(* Logix 5000 project; controller TFF vendor 1 type 14 code 107 rev 34.11; software revision 34.03; part 13 of 36 *)
(* tags used below, declared in another part *)
   AlarmAnalog : AlarmAnalog[50];   // Analog Alarm Array
   AlarmControl : AlarmControl;   // Alarm Control
   AlarmDeviation : AlarmDeviation[20];   // Control Loop Deviation Alarm Array
   AnalogPoint : AnalogInput[50];   // Analog Input Array
   CCPSystem : CCPSystem;   // CCP System Data
   ChartMark : ChartMark;   // Chart Mark
   Concentration : Concentration;
   ControlLoop : ControlLoop[20];   // Control Loop Array
   CriteriaFlag : CriteriaFlag;   // Criteria Flag used in CCP Recipe
   DCS : DCS;
   DerivedData : DerivedData;   // Derived data (user input and calculated values)
   Diafiltration : Diafiltration;
   DigitalPoint : DigitalPoint[150];   // Digital Point Array
   Drive : Drive[11];   // Drives Array
   FlowPath : FlowPath[64];   // Flow Path Array
   FlowPathControl : FlowPathControl;   // Flow Path Control
   FQ_Conc : ALIAS FOR Totalizer[0];   // Concentration Totalizer
   FQ_Diaf : ALIAS FOR Totalizer[1];   // DiafiltrationTotalizer
   LogVal : LoggedValue;   // Setpoints to be logged
   Membrane_Data : Membrane_Data;   // Membrane Data
   MiscBOOL : BOOL[64];   // Misc BOOL Values
   MiscDINT : DINT[32];   // Misc DINT Values
   MiscREAL : REAL[50];   // Misc Real Values
   Mixer : Mixer;   // Mixer config. structure
   Operation : Operation[6,251];   // Operation Table
   PCV001_Control : PCV_Control;   // PCV001 Control UDT
   PCV101_Control : PCV_Control;   // PCV101 Control UDT
   Phase : Phases[6];   // Phase Control Array
   Phase0 : ALIAS FOR Phase[0];   // Phase 0
   Phase1 : ALIAS FOR Phase[1];   // Phase 1
   Phase2 : ALIAS FOR Phase[2];   // Phase 2
   Phase3 : ALIAS FOR Phase[3];   // Phase 3
   Phase4 : ALIAS FOR Phase[4];   // Phase 4
   Phase5 : ALIAS FOR Phase[5];   // Phase 5
   PhaseTotalizer : PhaseTotalizer[18];   // Phase Totalizers Array
   Prompt : Prompt[7];   // Prompt Array
   Prompt0 : ALIAS FOR Prompt[0];   // Phase 0 Prompt
   Prompt1 : ALIAS FOR Prompt[1];   // Phase 1 Prompt
   Prompt2 : ALIAS FOR Prompt[2];   // Phase 2 Prompt
   Prompt3 : ALIAS FOR Prompt[3];   // Phase 3 Prompt
   Prompt4 : ALIAS FOR Prompt[4];   // Phase 4 Prompt
   Prompt5 : ALIAS FOR Prompt[5];   // Phase 5 Prompt
   PromptTimer : FBD_TIMER;   // Prompt Timer
   SRL001 : ALIAS FOR DigitalPoint[15];   // Tank Skid Remote / Standalone
   SysControl : SysControl;   // General system status and command
   Tank : TankManagement;   // Tank Management
   ThisSystem : SystemType;
   Timers : Timers[22];   // Timer Array
   Totalizer : Totalizers[20];   // Totalizers Array
   UserAlarm : UserAlarm;   // User Alarm (used in CCP Recipe)
   UserTotalizerManagement : UserTotalizerManagement;   // User Totalizer management
   Valve : Valve[100];   // Valve Array
   Y500A : ALIAS FOR DigitalOutput[11];   // Unlock Clamshell
   Y500B : ALIAS FOR DigitalOutput[12];   // Lock Clamshell
   Y501A : ALIAS FOR DigitalOutput[10];   // Unlock Door
   Y501B : ALIAS FOR DigitalOutput[9];   // Lock Door
   Y502A : ALIAS FOR DigitalOutput[13];   // Unlock Clamshell in Door
   Y502B : ALIAS FOR DigitalOutput[14];   // Lock Clamshell in Door
   Y503A : ALIAS FOR DigitalOutput[15];   // Connect Clamshell
   Y503B : ALIAS FOR DigitalOutput[16];   // Disconnect Clamshell

PROGRAM CCPSystem   (* main routine MainRoutine, fault routine FaultRoutine *)
VAR
   ActionCode : DINT := 1700011;   // Action Code
   ActionFlag : BOOL;   // Action Flag
   ActionProperty : DINT := 11;   // Action Property
   ActionStructure : DINT := 17;   // Action Data Structure
   ActionTag : DINT;   // Action Tag
   ActionValue : REAL := 1.0;   // Action Value
   AutoRunTimer : TIMER := (PRE := 5000);   // Auto Run Timer
   Boolean : DINT;   // Boolean Operator
        .1   // AND
        .0   // OR
   Branch : BOOL;   // Conditional Branch Flag
   BranchStep : DINT;   // Branch Step Number
   BufferStep : DINT := 60;   // Buffer Step
   Clear : BOOL;   // Clear Operation Table Flag
   Code : DINT := 3100002;   // Global Code
   CompleteTimer : TIMER := (PRE := 10000);   // Operation Complete Timer
   Criteria1BoolValue : BOOL;   // Criteria 1 Discrete Value
   Criteria1Code : DINT := 1100602;   // Criteria 1 Code
   Criteria1Met : BOOL := 1;   // Criteria 1 Met
   Criteria1Operator : DINT := 1;   // Criteria 1 Operator
        .0   // >=
        .1   // <=
        .2   // =
   Criteria1Property : DINT := 2;   // Criteria 1 Property
   Criteria1RealValue : REAL := 2.0;   // Criteria 1 Real Value
   Criteria1Structure : DINT := 11;   // Criteria 1 Data Structure
   Criteria1Tag : DINT := 6;   // Criteria 1 Tag
   Criteria1Type : BOOL;   // Criteria 1 Type 0=Real, 1=Boolean
   Criteria1Value : REAL := 2.0;   // Criteria 1 Value
   Criteria2BoolValue : BOOL := 1;   // Criteria 2 Discrete Value
   Criteria2Code : DINT;   // Criteria 2 Code
   Criteria2Met : BOOL := 1;   // Criteria 2 Met
   Criteria2Operator : DINT;   // Criteria 2 Operator
        .0   // >=
        .1   // <=
        .2   // =
   Criteria2Property : DINT := 3;   // Criteria 2 Property
   Criteria2RealValue : REAL := 6.0;   // Criteria 2 Real Value
   Criteria2Structure : DINT;   // Criteria 2 Data Structure
   Criteria2Tag : DINT;   // Criteria 2 Tag
   Criteria2Type : BOOL;   // Criteria 2 Type 0=Real, 1=Boolean
   Criteria2Value : REAL;   // Criteria 2 Value
   CriteriaMet : BOOL := 1;   // Criteria Met
   DateTime : DINT[7] := ([0] := 2026, [1] := 7, [2] := 24, [3] := 11, [4] := 48, [5] := 55, [6] := 561276);   // Date and Time
   DownloadONS : BOOL;
   EnableStep : BOOL;   // Step Action Enabled
   ErrorCheck : BOOL;   // Error Check Flag
   ErrorCheckONS : BOOL := 1;   // Error Check One-Shot
   Index : DINT := 585;   // Index
   LastStep : DINT := 59;   // Last Step
   NextStep : DINT := 61;   // Next Step
   PendingStep : DINT := 61;   // Current Step
   Phase0StopONS : BOOL;
   PhaseClear : BOOL;   // Phase Clear
   PhaseClearNumber : DINT := 6;   // Phase Clear Number
   PhaseNumber : DINT := 6;   // Phase FOR NEXT Index
   Pointer : DINT := 85;   // Pointer
   PreRunLog : BOOL;   // Log Pre Run Set Points
   Property : DINT := 2;   // Case Property
   ResumeDownloadFromHOLD : BOOL;
   Run : BOOL;   // Operation Run Status
   RunONS : BOOL;   // Run Command One-Shot
   sAction : STRING10 := '1700011';   // Action Code String
   sActionProperty : STRING4 := '11';   // Action Property String
   sActionStructure : STRING4 := '17';   // Action Data Structure String
   sActionTag : STRING4 := '000';   // Action Tag String
   sBufferEvents : STRING50 := '07242026,11:31:58.3,305006,1.00000000,';   // Buffer Events String
   sCode : STRING10 := '1900011';   // Global code String
   sColon : STRING4 := ':';   // Colon separator String
   sComma : STRING4 := ',';   // Comma String
   sCriteria1 : STRING10 := '1100602';   // Criteria 1 Code String
   sCriteria1Property : STRING4 := '02';   // Criteria 1 Property String
   sCriteria1Structure : STRING4 := '11';   // Criteria 1 Data Structure String
   sCriteria1Tag : STRING4 := '006';   // Criteria 1 Tag String
   sCriteria2 : STRING10 := '800003';   // Criteria 2 Code String
   sCriteria2Property : STRING4 := '03';   // Criteria 2 Property String
   sCriteria2Structure : STRING4 := '8';   // Criteria 2 Data Structure String
   sCriteria2Tag : STRING4 := '000';   // Criteria 2 Tag String
   sDateTime : STRING25 := '07242026,11:48:55.6,';   // Date and Time String
   sPeriod : STRING4 := '.';   // Timer separator String
   sProperty : STRING4 := '02';   // Property String
   sStructure : STRING4 := '9';   // Structure String
   sTag : STRING4 := '000';   // Tag String
   sTemp : STRING50 := '8';   // Temp String
   Structure : DINT := 1;   // Structure code
   sZero : STRING4 := '0';   // Zero String
   Tag : DINT;   // Tag value
   TempEvents : DINT := 50;   // Temp Register
   TempSteps : DINT := 26;
   Tenths : DINT := 8;   // Thents (Date and Time management)
   ThisStep : DINT := 21;   // This Step (Error management)
   Value : REAL;   // Temp Value
END_VAR

ROUTINE Action   (* structured text *)
// Operation Action Routine
   (* =======================================================================
   	Operation Action : Get the current action code and perform action based on information extraction
   
   	List of treatments
   		- Get current action code
   		- Extract informations based on action code
   		- Navigate through the action categories to perform action
   		- Jump to BufferSteps routine and update step numbers
   
   -----------------------------------------------------------------------------------------------------------------------------------------------------
   	History
   		2019-AUG-13 - ACTEMIUM - B. Roch - Initial version for Candidate Release 3.00.00.00.a
   		2019-SEP-09 - ACTEMIUM - Q. Spindler - Modifications for Candidate Release 3.00.00.00.c
   					- Fix Clamchell Actions YA502A, YA502B, YA503A, and YA503B
   		2022-FEB-14 - Davidson - Ch.Arbogast - Modifications for Candidate Release 3.02.00.00.a
   			- On 8 Case 1 + 2, add Reset of ResponseOK, YES, and NO on prompt action
   			- Case 30, add DCS Actions for pumps setpoints, PCV setpoints, Mixer setpoints, Protein Conc., Holdup + Diaf Volume, membrane area + density
   =========================================================================*)
   
   
   (* Get current action code
   =========================================================================*)
   (*Get the pending step Action Code and Action Value from the operation array*)
   ActionCode := Operation[PhaseNumber,PendingStep].Action;
   ActionValue := Operation[PhaseNumber,PendingStep].ActionValue;
   
   (* Extract informations based on action code
   =========================================================================*)
   (*Extract the Structure, Tag and Property values from the action code. The action code is
   in the format SSTTTPP  SS is Structure Element, TTT is action TagElement i.e ControlLoop[TTT].Enable
   PP Action Property Number in secound Case below.*)
   
   IF ActionCode <> 0 THEN;
   	DTOS (ActionCode, sAction);
   	IF sAction.LEN = 7 THEN;
   		MID (sAction, 2, 1, sActionStructure);
   		MID (sAction, 3, 3, sActionTag);
   		MID (sAction, 2, 6, sActionProperty);
   	ELSIF sAction.LEN = 6 THEN;
   		MID (sAction, 1, 1, sActionStructure);
   		MID (sAction, 3, 2, sActionTag);
   		MID (sAction, 2, 5, sActionProperty);
   	ELSIF sAction.LEN = 5 THEN;
   		(* Ignore if code length is not 6 or 7 *)
   		DTOS(0,sActionStructure);
   	ELSE;
   		CCPSystem.Error := 7;
   	END_IF;
   	STOD (sActionStructure, ActionStructure);
   	STOD (sActionTag, ActionTag);
   	STOD (sActionProperty, ActionProperty);
   ELSE;
   	ActionStructure := 0;
   END_IF;
   
   (* Navigate through the action categories to perform action
   =========================================================================*)
   CASE ActionStructure OF
   	0:	; (*No Action)*)
   	1: 	CASE	ActionProperty OF (*Analog Alarms*)
   			1:	IF NOT ErrorCheck THEN; IF ActionValue = 0 THEN AlarmAnalog[ActionTag].Override := 0; ELSE AlarmAnalog[ActionTag].Override := 1; END_IF; END_IF;
   			2:	IF NOT ErrorCheck THEN; AlarmAnalog[ActionTag].LOLO := ActionValue; END_IF;
   			3:	IF NOT ErrorCheck THEN; AlarmAnalog[ActionTag].LO := ActionValue; END_IF;
   			4:	IF NOT ErrorCheck THEN; AlarmAnalog[ActionTag].HI := ActionValue; END_IF;
   			5:	IF NOT ErrorCheck THEN; AlarmAnalog[ActionTag].HIHI := ActionValue; END_IF;
   		ELSE 	CCPSystem.Error := 7;
   		END_CASE;
   	2:	CASE	ActionProperty OF (*Deviation Alarms*)
   			1:	IF NOT ErrorCheck THEN; IF ActionValue = 0 THEN AlarmDeviation[ActionTag].Override := 0; ELSE AlarmDeviation[ActionTag].Override := 1; END_IF; END_IF;
   			4:	IF NOT ErrorCheck THEN; AlarmDeviation[ActionTag].HI := ActionValue; END_IF;
   			5:	IF NOT ErrorCheck THEN; AlarmDeviation[ActionTag].HIHI := ActionValue; END_IF;
   		ELSE 	CCPSystem.Error := 7;
   		END_CASE;
   	3:	CASE	ActionProperty OF (*Digital Alarms*)
   			1:	IF NOT ErrorCheck THEN; IF ActionValue = 0 THEN DigitalPoint[ActionTag].Override := 0; ELSE DigitalPoint[ActionTag].Override := 1; END_IF; END_IF;
   		ELSE 	CCPSystem.Error := 7;
   		END_CASE;
   	5:	CASE	ActionProperty OF (*Control Loops*)
   			1:	IF NOT ErrorCheck THEN; IF ActionValue = 0 THEN ControlLoop[ActionTag].Manual := 0; ELSE ControlLoop[ActionTag].Manual := 1; END_IF; END_IF;
   			2:	IF NOT ErrorCheck THEN; IF ActionValue = 0 THEN ControlLoop[ActionTag].Auto1 := 0; ELSE ControlLoop[ActionTag].Auto1 := 1; END_IF; END_IF;
   			3:	IF NOT ErrorCheck THEN; IF ActionValue = 0 THEN ControlLoop[ActionTag].Auto2 := 0; ELSE ControlLoop[ActionTag].Auto2 := 1; END_IF; END_IF;
   			4:	IF NOT ErrorCheck THEN; IF ActionValue = 0 THEN ControlLoop[ActionTag].Auto3 := 0; ELSE ControlLoop[ActionTag].Auto3 := 1; END_IF; END_IF;
   			5:	IF NOT ErrorCheck THEN; IF ActionValue = 0 THEN ControlLoop[ActionTag].Auto4 := 0; ELSE ControlLoop[ActionTag].Auto4 := 1; END_IF; END_IF;
   			6:	IF NOT ErrorCheck THEN; ControlLoop[ActionTag].SPManual := ActionValue; END_IF;
   			7:	IF NOT ErrorCheck THEN; ControlLoop[ActionTag].SPAuto1 := ActionValue; END_IF;
   			8:	IF NOT ErrorCheck THEN; ControlLoop[ActionTag].SPAuto2 := ActionValue; END_IF;
   			9:	IF NOT ErrorCheck THEN; ControlLoop[ActionTag].SPAuto3 := ActionValue; END_IF;
   			10:	IF NOT ErrorCheck THEN; ControlLoop[ActionTag].SPAuto4 := ActionValue; END_IF;
   			11:	IF NOT ErrorCheck THEN; ControlLoop[ActionTag].RampRate := ActionValue; END_IF;
   			12:	IF NOT ErrorCheck THEN; ControlLoop[ActionTag].Deadband := ActionValue; END_IF;
   			13:	IF NOT ErrorCheck THEN; ControlLoop[ActionTag].StableTime := ActionValue; END_IF;
   			14:	IF NOT ErrorCheck THEN; ControlLoop[ActionTag].KP[0] := ActionValue; END_IF;
   			15:	IF NOT ErrorCheck THEN; ControlLoop[ActionTag].KI[0] := ActionValue; END_IF;
   			16:	IF NOT ErrorCheck THEN; ControlLoop[ActionTag].KD[0] := ActionValue; END_IF;
   			17:	IF NOT ErrorCheck THEN; ControlLoop[ActionTag].DB[0] := ActionValue; END_IF;
   			18:	IF NOT ErrorCheck THEN; ControlLoop[ActionTag].KP[1] := ActionValue; END_IF;
   			19:	IF NOT ErrorCheck THEN; ControlLoop[ActionTag].KI[1] := ActionValue; END_IF;
   			20:	IF NOT ErrorCheck THEN; ControlLoop[ActionTag].KD[1] := ActionValue; END_IF;
   			21: IF NOT ErrorCheck THEN; ControlLoop[ActionTag].DB[1] := ActionValue; END_IF;
   			22: IF NOT ErrorCheck THEN; ControlLoop[ActionTag].KP[2] := ActionValue; END_IF;
   			23:	IF NOT ErrorCheck THEN; ControlLoop[ActionTag].KI[2] := ActionValue; END_IF;
   			24:	IF NOT ErrorCheck THEN; ControlLoop[ActionTag].KD[2] := ActionValue; END_IF;
   			25:	IF NOT ErrorCheck THEN; ControlLoop[ActionTag].DB[2] := ActionValue; END_IF;
   		ELSE 	CCPSystem.Error := 7;
   		END_CASE;
   	7:	CASE	ActionProperty OF (*Phase Control*)
   			1:	IF NOT ErrorCheck THEN; IF ActionValue = 0 THEN Phase[ActionTag].Run := 0; ELSE Phase[ActionTag].Run := 1; END_IF; END_IF;
   			2:	IF NOT ErrorCheck THEN; IF ActionValue = 0 THEN Phase[ActionTag].Stop := 0; ELSE Phase[ActionTag].Stop := 1; END_IF; END_IF;
   			3:	IF NOT ErrorCheck THEN; IF ActionValue = 0 THEN Phase[ActionTag].Hold := 0; ELSE Phase[ActionTag].Hold := 1; END_IF; END_IF;
   			4:	IF NOT ErrorCheck THEN; IF ActionValue = 0 THEN Phase[ActionTag].Pause := 0; ELSE Phase[ActionTag].Pause := 1; END_IF; END_IF;
   			5:	IF NOT ErrorCheck THEN;
   				Phase[PhaseNumber].JumpPLC := 1; (*Conditional Branch*)
   				Phase[PhaseNumber].ActualStep := BranchStep;
   				END_IF;
   		ELSE 	CCPSystem.Error := 7;
   		END_CASE;
   	8:	CASE	ActionProperty OF (*Prompts*)
   			(*Prompts OK*)
   			1:	IF NOT ErrorCheck THEN;
   					(*Delay to Prompts to allow back to back*)
   					TONR(PromptTimer);
   					PromptTimer.EN := 1;
   					PromptTimer.PRE := 1000;
   					while PromptTimer.TT and Prompt[PhaseNumber].PromptOK   do;
   					end_while;
   				Prompt[PhaseNumber].PromptYesNO := 0;
   				Prompt[PhaseNumber].PromptOK := 1;
   				Prompt[PhaseNumber].ResponseOK := 0;
   				Prompt[PhaseNumber].Step := PendingStep;
   				Prompt[PhaseNumber].Flag := 1;
   				Prompt[PhaseNumber].Pending := 1;
   				Prompt[PhaseNumber].Value := ActionValue; (*PV+*)
   				END_IF;
   			(*Prompts YesNo*)
   			2:	IF NOT ErrorCheck THEN;
   					(*Delay to Prompts to allow back to back*)
   					TONR(PromptTimer);
   					PromptTimer.EN := 1;
   					PromptTimer.PRE := 1000;
   					while PromptTimer.TT and Prompt[PhaseNumber].PromptYesNO do;
   					end_while;
   				Prompt[PhaseNumber].PromptOK := 0;
   				Prompt[PhaseNumber].PromptYesNO := 1;
   				Prompt[PhaseNumber].ResponseNo := 0;
   				Prompt[PhaseNumber].ResponseYes := 0;
   				Prompt[PhaseNumber].Step := PendingStep;
   				Prompt[PhaseNumber].Flag := 1;
   				Prompt[PhaseNumber].Pending := 1;
   				END_IF;
   			3:	IF NOT ErrorCheck THEN;
   				Prompt[PhaseNumber].Flag := 1;
   				Prompt[PhaseNumber].Step := PendingStep;
   				END_IF;
   		ELSE 	CCPSystem.Error := 7;
   		END_CASE;
   	9:	CASE	ActionProperty OF (*Pumps*)
   			1:	IF NOT ErrorCheck THEN; IF ActionValue = 0 THEN Drive[ActionTag].AutoCommand := 0; ELSE Drive[ActionTag].AutoCommand := 1; END_IF; END_IF;
   			2:	IF NOT ErrorCheck THEN; IF ActionValue = 0 THEN Drive[ActionTag].Direction := 0; ELSE Drive[ActionTag].Direction := 1; END_IF; END_IF;
   		ELSE 	CCPSystem.Error := 7;
   		END_CASE;
   	11:	CASE	ActionProperty OF (*Timers*)
   			3:	IF NOT ErrorCheck THEN; IF ActionValue = 0 THEN Timers[ActionTag].Enable := 0; ELSE Timers[ActionTag].Enable := 1; END_IF; END_IF;
   			4:	IF NOT ErrorCheck THEN; IF ActionValue = 0 THEN Timers[ActionTag].Reset := 0; ELSE Timers[ActionTag].Reset := 1; END_IF; END_IF;
   		ELSE 	CCPSystem.Error := 7;
   		END_CASE;
   	12:	CASE	ActionProperty OF (*Totalizers*)
   			6:	IF NOT ErrorCheck THEN; IF ActionValue = 0 THEN Totalizer[0].Enable := 0; ELSE Totalizer[0].Enable := 1; END_IF; END_IF;
   			7:	IF NOT ErrorCheck THEN; Totalizer[0].Reset := 1; END_IF;
   			8:	IF NOT ErrorCheck THEN; IF ActionValue = 0 THEN Totalizer[1].Enable := 0; ELSE Totalizer[1].Enable := 1; END_IF; END_IF;
   			9:	IF NOT ErrorCheck THEN; Totalizer[1].Reset := 1; END_IF;
   		ELSE 	CCPSystem.Error := 7;
   		END_CASE;
   	13:	CASE	ActionProperty OF (*Valves*)
   			1:	IF NOT ErrorCheck THEN; IF ActionValue = 0 THEN Valve[ActionTag].Auto := 0; ELSE Valve[ActionTag].Auto := 1; END_IF; END_IF;
   		ELSE 	CCPSystem.Error := 7;
   		END_CASE;
   	14:	CASE	ActionProperty OF (*Mixer*)
   			1:	IF NOT ErrorCheck THEN; IF ActionValue = 0 THEN Mixer.Mode := 0; ELSE Mixer.Mode := 1; END_IF; END_IF;
   			2:	IF NOT ErrorCheck THEN; Mixer.SPManual := ActionValue; END_IF;
   			3:	IF NOT ErrorCheck THEN; Mixer.SPAutoMin := ActionValue; END_IF;
   			4:	IF NOT ErrorCheck THEN; Mixer.SPAutoMax := ActionValue; END_IF;
   			5:	IF NOT ErrorCheck THEN; Mixer.LevelMin := ActionValue; END_IF;
   			6:	IF NOT ErrorCheck THEN; Mixer.LevelMax := ActionValue; END_IF;
   		ELSE 	CCPSystem.Error := 7;
   		END_CASE;
   	15:	CASE	ActionProperty OF (*Misc.*)
   			1:	IF NOT ErrorCheck THEN; IF ActionValue = 0 THEN MiscBOOL[ActionTag] := 0; ELSE MiscBOOL[ActionTag] := 1; END_IF; END_IF;
   			2:	IF NOT ErrorCheck THEN; MiscDINT[ActionTag] := ActionValue; END_IF;
   			3:	IF NOT ErrorCheck THEN; MiscREAL[ActionTag] := ActionValue; END_IF;
   		ELSE 	CCPSystem.Error := 7;
   		END_CASE;
   	16:	CASE	ActionProperty OF (*Alarm Control*)
   			1:	IF NOT ErrorCheck THEN; AlarmControl.EnableAllIn := 1; END_IF;
   			2:	IF NOT ErrorCheck THEN; AlarmControl.DisableAllIn := 1; END_IF;
   			6:	IF NOT ErrorCheck THEN; AlarmControl.EnableAllAnaSigIn := 1; END_IF;
   			7:	IF NOT ErrorCheck THEN; AlarmControl.DisableAllAnaSigIn := 1; END_IF;
   		ELSE 	CCPSystem.Error := 7;
   		END_CASE;
   	17:	CASE	ActionProperty OF (*Miscellaneous*)
   			1:	IF NOT ErrorCheck THEN; SysControl.DefaultIn := 1; END_IF;
   			2:	IF NOT ErrorCheck THEN; ChartMark.In := 1; END_IF;
   			3:	IF NOT ErrorCheck THEN; SysControl.AllAutoIn := 1; END_IF;
   			4:	IF NOT ErrorCheck THEN; UserTotalizerManagement.LogUserIn := 1; END_IF;
   			5:	IF NOT ErrorCheck THEN; IF ActionValue = 0 THEN UserTotalizerManagement.StartUser := 0; ELSE UserTotalizerManagement.StartUser := 1; END_IF; END_IF;
   			6:	IF NOT ErrorCheck THEN; UserTotalizerManagement.ResetUserIn:= 1; END_IF;
   			7:	IF NOT ErrorCheck THEN; Tank.Feed_Bag_Tare := 1; END_IF;
   			8:	IF NOT ErrorCheck THEN; Tank.Filtrate_Bag_Tare := 1; END_IF;
   			9:	IF NOT ErrorCheck THEN; SysControl.UV_Auto_Zero_Cmd := 1; END_IF;
   			11:	IF NOT ErrorCheck THEN; IF ActionValue = 0 THEN CCPSystem.DefaultOnComplete := 0; ELSE CCPSystem.DefaultOnComplete := 1; END_IF; END_IF;
   			12:	IF NOT ErrorCheck THEN; UserAlarm.NonCritical1 := 1; END_IF;
   			13:	IF NOT ErrorCheck THEN; UserAlarm.Critical1 := 1; END_IF;
   			14:	IF NOT ErrorCheck THEN; UserAlarm.NonCritical2 := 1; END_IF;
   			15:	IF NOT ErrorCheck THEN; UserAlarm.Critical2 := 1; END_IF;
   		ELSE 	CCPSystem.Error := 7;
   		END_CASE;
   	18:	CASE	ActionProperty OF (*Criteria Flag*)
   			1:	IF NOT ErrorCheck THEN; IF ActionValue = 0 THEN CriteriaFlag.Flag1 := 0; ELSE CriteriaFlag.Flag1 := 1; END_IF; END_IF;
   			2:	IF NOT ErrorCheck THEN; IF ActionValue = 0 THEN CriteriaFlag.Flag2 := 0; ELSE CriteriaFlag.Flag2 := 1; END_IF; END_IF;
   			3:	IF NOT ErrorCheck THEN; IF ActionValue = 0 THEN CriteriaFlag.Flag3 := 0; ELSE CriteriaFlag.Flag3 := 1; END_IF; END_IF;
   			4:	IF NOT ErrorCheck THEN; IF ActionValue = 0 THEN CriteriaFlag.Flag4 := 0; ELSE CriteriaFlag.Flag4 := 1; END_IF; END_IF;
   			5:	IF NOT ErrorCheck THEN; IF ActionValue = 0 THEN CriteriaFlag.Flag5 := 0; ELSE CriteriaFlag.Flag5 := 1; END_IF; END_IF;
   		ELSE 	CCPSystem.Error := 7;
   		END_CASE;
   	19:	CASE	ActionProperty OF (*Concentration*)
   			1:	IF NOT ErrorCheck THEN; IF ActionValue = 0 THEN FQ_Conc.Enable := 0; ELSE FQ_Conc.Enable := 1; END_IF; END_IF;
   			2:	IF NOT ErrorCheck THEN; FQ_Conc.Reset:= 1; END_IF;
   			3:	IF NOT ErrorCheck THEN; Concentration.LogConcIn := 1; END_IF;
   			4:	IF NOT ErrorCheck THEN; Concentration.Conc_Init := ActionValue; END_IF;
   			5:	IF NOT ErrorCheck THEN; Concentration.Conc_Final := ActionValue; END_IF;
   			6:	IF NOT ErrorCheck THEN; Concentration.Conc_Final_Volume := ActionValue; END_IF;
   			7:	IF NOT ErrorCheck THEN; DerivedData.HOLDUP := ActionValue; END_IF;
   		ELSE 	CCPSystem.Error := 7;
   		END_CASE;
   	20:	CASE	ActionProperty OF (*Diafiltration*)
   			1:	IF NOT ErrorCheck THEN; IF ActionValue = 0 THEN FQ_Diaf.Enable := 0; ELSE FQ_Diaf.Enable := 1; END_IF; END_IF;
   			2:	IF NOT ErrorCheck THEN; FQ_Diaf.Reset:= 1; END_IF;
   			3:	IF NOT ErrorCheck THEN; Diafiltration.LogDiafIn := 1; END_IF;
   			4:	IF NOT ErrorCheck THEN; Diafiltration.Snap := 1; END_IF;
   			5:	IF NOT ErrorCheck THEN; Diafiltration.Diaf_Init := ActionValue; END_IF;
   			6:	IF NOT ErrorCheck THEN; Diafiltration.Diaf_Final_Volume := ActionValue; END_IF;
   		ELSE 	CCPSystem.Error := 7;
   		END_CASE;
   	21:	CASE	ActionProperty OF (*Membrane Data*)
   			1:	IF NOT ErrorCheck THEN; Membrane_Data.Area := ActionValue; END_IF;
   			2:	IF NOT ErrorCheck THEN; Membrane_Data.Density := ActionValue; END_IF;
   		ELSE 	CCPSystem.Error := 7;
   		END_CASE;
   	23:	CASE	ActionProperty OF (*PCV Control*)
   			1:	IF NOT ErrorCheck THEN; PCV001_Control.FullOpen := 1; END_IF;
   			2:	IF NOT ErrorCheck THEN; PCV001_Control.FullClose := 1; END_IF;
   			3:	IF NOT ErrorCheck THEN; PCV101_Control.FullOpen := 1; END_IF;
   			4:	IF NOT ErrorCheck THEN; PCV101_Control.FullClose := 1; END_IF;
   		ELSE 	CCPSystem.Error := 7;
   		END_CASE;
   	24:	CASE	Property OF (*Event value.*)
   			1:	IF NOT ErrorCheck THEN; LogVal.Value[Tag] := ActionValue; END_IF;
   		ELSE 	CCPSystem.Error := 7;
   		END_CASE;
   	25:	CASE	ActionProperty OF (*Flow Paths*)
   			1:	IF NOT ErrorCheck THEN; IF ActionValue = 0 THEN FlowPath[ActionTag].Command := 0; ELSE FlowPath[ActionTag].Command := 1; END_IF; END_IF;
   			2:	IF NOT ErrorCheck THEN; IF ActionValue = 0 THEN FlowPathControl.FlushMode_Enabled := 0; ELSE FlowPathControl.FlushMode_Enabled := 1; END_IF; END_IF;
   			3:	IF NOT ErrorCheck THEN; IF ActionValue = 0 THEN FlowPathControl.DrainMode_Enabled := 0; ELSE FlowPathControl.DrainMode_Enabled := 1; END_IF; END_IF;
   		ELSE 	CCPSystem.Error := 7;
   		END_CASE;
   	26:	CASE	ActionProperty OF (*Clamshell*)
   			1:	IF NOT ErrorCheck THEN; IF ActionValue = 0 THEN Y500A := 0; ELSE Y500A := 1; END_IF; END_IF;
   			2:	IF NOT ErrorCheck THEN; IF ActionValue = 0 THEN Y500B := 0; ELSE Y500B := 1; END_IF; END_IF;
   			3:	IF NOT ErrorCheck THEN; IF ActionValue = 0 THEN Y501A := 0; ELSE Y501A := 1; END_IF; END_IF;
   			4:	IF NOT ErrorCheck THEN; IF ActionValue = 0 THEN Y501B := 0; ELSE Y501B := 1; END_IF; END_IF;
   			5:	IF NOT ErrorCheck THEN; IF ActionValue = 0 THEN Y502A := 0; ELSE Y502A := 1; END_IF; END_IF;
   			6:	IF NOT ErrorCheck THEN; IF ActionValue = 0 THEN Y502B := 0; ELSE Y502B := 1; END_IF; END_IF;
   			7:	IF NOT ErrorCheck THEN; IF ActionValue = 0 THEN Y503A := 0; ELSE Y503A := 1; END_IF; END_IF;
   			8:	IF NOT ErrorCheck THEN; IF ActionValue = 0 THEN Y503B := 0; ELSE Y503B := 1; END_IF; END_IF;
   		ELSE 	CCPSystem.Error := 7;
   		END_CASE;
   
   		30:	CASE	ActionProperty OF (*DCS*)
   			0:	IF NOT ErrorCheck THEN; ControlLoop[1].SPManual := DCS.ActionsParameters.Feed_Pump_Speed_Setpoint[ActionTag]; END_IF;
   			1:	IF NOT ErrorCheck THEN; ControlLoop[1].SPAuto1 := DCS.ActionsParameters.Feed_Pump_Flow_Setpoint[ActionTag]; END_IF;
   			2:	IF NOT ErrorCheck THEN; ControlLoop[1].SPAuto2 := DCS.ActionsParameters.Feed_Pump_DP_Setpoint[ActionTag]; END_IF;
   			3:	IF NOT ErrorCheck THEN; ControlLoop[2].SPManual := DCS.ActionsParameters.Level_Pump_Speed_Setpoint[ActionTag]; END_IF;
   			4:	IF NOT ErrorCheck THEN; ControlLoop[2].SPAuto1 := DCS.ActionsParameters.Level_Pump_Level_Setpoint[ActionTag]; END_IF;
   			6:	IF NOT ErrorCheck THEN; ControlLoop[3].SPManual := DCS.ActionsParameters.PCV001_Retentate_Position_Setpoint[ActionTag]; END_IF;
   			7:	IF NOT ErrorCheck THEN; ControlLoop[3].SPAuto1 := DCS.ActionsParameters.PCV001_Retentate_Pressure_Setpoint[ActionTag]; END_IF;
   			8:	IF NOT ErrorCheck THEN; ControlLoop[3].SPAuto2 := DCS.ActionsParameters.PCV001_Retentate_TMP_Setpoint[ActionTag]; END_IF;
   			9:	IF NOT ErrorCheck THEN; ControlLoop[5].SPManual := DCS.ActionsParameters.PCV101_Filtrate_Position_Setpoint[ActionTag]; END_IF;
   			10:	IF NOT ErrorCheck THEN; ControlLoop[5].SPAuto1 := DCS.ActionsParameters.PCV101_Filtrate_Flow_Setpoint[ActionTag]; END_IF;
   			11:	IF NOT ErrorCheck THEN; ControlLoop[5].SPAuto2 := DCS.ActionsParameters.PCV101_Filtrate_TMP_Setpoint[ActionTag]; END_IF;
   			12:	IF NOT ErrorCheck THEN; Mixer.SPManual := DCS.ActionsParameters.Mixer_Speed_Setpoint[ActionTag]; END_IF;
   			13:	IF NOT ErrorCheck THEN; Mixer.SPAutoMin := DCS.ActionsParameters.Mixer_Auto_Min_Setpoint[ActionTag]; END_IF;
   			14:	IF NOT ErrorCheck THEN; Mixer.SPAutoMax := DCS.ActionsParameters.Mixer_Auto_Max_Setpoint[ActionTag]; END_IF;
   			15:	IF NOT ErrorCheck THEN; Concentration.Conc_Init := DCS.ActionsParameters.Init_Protein_Conc[ActionTag]; END_IF;
   			16:	IF NOT ErrorCheck THEN; Concentration.Conc_Final := DCS.ActionsParameters.Final_Protein_Conc[ActionTag]; END_IF;
   			17:	IF NOT ErrorCheck THEN; Concentration.Conc_Final_Volume := DCS.ActionsParameters.Final_Protein_Volume[ActionTag]; END_IF;
   			18:	IF NOT ErrorCheck THEN; DerivedData.HOLDUP := DCS.ActionsParameters.Holdup_Volume[ActionTag]; END_IF;
   			19:	IF NOT ErrorCheck THEN; Diafiltration.Diaf_Init := DCS.ActionsParameters.Init_Diaf_Volume[ActionTag]; END_IF;
   			20:	IF NOT ErrorCheck THEN; Diafiltration.Diaf_Final_Volume := DCS.ActionsParameters.Final_Diaf_Volume[ActionTag]; END_IF;
   			21:	IF NOT ErrorCheck THEN; Membrane_Data.Area := DCS.ActionsParameters.Membrane_Area[ActionTag]; END_IF;
   			22:	IF NOT ErrorCheck THEN; Membrane_Data.Density := DCS.ActionsParameters.Membrane_Density[ActionTag]; END_IF;
   		ELSE 	CCPSystem.Error := 7;
   		END_CASE;
   ELSE 	CCPSystem.Error := 7;
   END_CASE;
   
   (* Jump to BufferSteps routine and update step numbers
   =========================================================================*)
   IF NOT ErrorCheck THEN;
   	JSR (BufferSteps);
   	IF NOT Phase[PhaseNumber].JumpPLC THEN;
   		(*Update Actual step, pending step and jump step number*)
   		Phase[PhaseNumber].ActualStep := PendingStep + 1;
   		PendingStep := PendingStep + 1;
   		Phase[PhaseNumber].JumpStep := PendingStep + 1;
   	END_IF;
   END_IF;
END_ROUTINE

ROUTINE Branch   (* structured text *)
// Branch to Label Routine
   (* =======================================================================
   	Branch : Conditionnal branch management
   
   	List of treatments
   		- Get current action code
   		- Extract informations based on action code
   		- Jump to label and Jump Step processing
   
   -----------------------------------------------------------------------------------------------------------------------------------------------------
   	History
   		2019-AUG-13 - ACTEMIUM - B. Roch - Initial version for Candidate Release 3.00.00.00.a
   =========================================================================*)
   
   
   (* Get current action code
   =========================================================================*)
   (*Get the pending step Action Code and Action Value from the operation array*)
   ActionCode := Operation[PhaseNumber,PendingStep].Action;
   ActionValue := Operation[PhaseNumber,PendingStep].ActionValue;
   
   (* Extract informations based on action code
   =========================================================================*)
   (*Extract the Structure, Tag and Property values from the action code. The action code is
   in the format SSTTTPP*)
   IF ActionCode <> 0 THEN;
   	DTOS (ActionCode, sAction);
   	IF sAction.LEN = 7 THEN;
   		MID (sAction, 2, 1, sActionStructure);
   		MID (sAction, 3, 3, sActionTag);
   		MID (sAction, 2, 6, sActionProperty);
   	ELSIF sAction.LEN = 6 THEN;
   		MID (sAction, 1, 1, sActionStructure);
   		MID (sAction, 3, 2, sActionTag);
   		MID (sAction, 2, 5, sActionProperty);
   	END_IF;
   	STOD (sActionStructure, ActionStructure);
   	STOD (sActionTag, ActionTag);
   	STOD (sActionProperty, ActionProperty);
   ELSE;
   	ActionStructure := 0;
   	ActionProperty := 0;
   END_IF;
   
   (* Jump to label and Jump Step processing
   =========================================================================*)
   (*Check to determine if action is a conditional branch, Structure=7 and Property=5*)
   BranchStep := 0;
   Phase[PhaseNumber].Label := 0;
   IF ActionStructure = 7 AND ActionProperty = 5  AND NOT Prompt[PhaseNumber].Pending THEN;
   	IF CriteriaMet THEN;
   		FOR BranchStep := 1 TO 250 DO;
   		(*If Jump to label action exist copy the label value in corresponding Phase label*)
   			IF Operation[PhaseNumber, BranchStep].Label = ActionValue THEN;
   				Phase[PhaseNumber].Label := ActionValue;
   				EXIT;
   			END_IF;
   		END_FOR;
   	ELSE;
   		(*Jump to BufferSteps routine and update Actual step number*)
   		JSR (BufferSteps);
   		Phase[PhaseNumber].ActualStep := (PendingStep + 1);
   	END_IF;
   
   ELSIF Phase[PhaseNumber].JumpPLC THEN;
   	FOR BranchStep := 1 TO 250 DO;
   		IF Operation[PhaseNumber, BranchStep].Step = Phase[PhaseNumber].JumpStep THEN;
   			Phase[PhaseNumber].ActualStep := BranchStep;
   			EXIT;
   		END_IF;
   	END_FOR;
   END_IF;
   
END_ROUTINE

ROUTINE BufferEvents   (* structured text *)
// Event Log Buffer Routine
   (* =======================================================================
   	Buffer Events : This routine scans all event code values defined in the event array downloaded by CCP6
   					If the value of the tag referenced by the code has changed from the last scan,the time stamp,
   					action code and new/old values are written to the buffer.
   					The buffer pointer used by CCP6 is updated after scanning all tags
   
   	Warning :		This code should not be modified without a control of change impact on the Recipe download check procedure of CCPRuntime.exe
   
   	List of treatments
   		- Get current action code
   		- Extract informations based on event code
   		- Navigate through the event categories
   		- Log Pre-run values
   		- Build event contents
   		- Reset flag and pointer
   
   -----------------------------------------------------------------------------------------------------------------------------------------------------
   	History
   		2019-AUG-13 - ACTEMIUM - B. Roch - Initial version for Candidate Release 3.00.00.00.a
   		2022-FEB-14 - Davidson - Ch.Arbogast - Modifications for Candidate Release 3.02.00.00.a
   			- Change resetting of sStructure in case of wrong code length by DTOS function :
   			  On Ignore if code length is not 6 or 7, replace "sStructure.DATA[0] := sZero.DATA[0]"
   			  by "DTOS (0, sStructure)"
   			- Case 17, add Tamk Skid Remote / standalone Event
   			- Case 30, add DCS Actions for Mixing pumps setpoints, primary and secondary conductivity, Deadbands, and stable times
   			- Case 31: add DCS Criteria
   =========================================================================*)
   
   
   (* Get the current pointer value
   =========================================================================*)
   STOD (CCPSystem.BufferEvents[0], Pointer);
   
   (* Extract informations based on event code
   =========================================================================*)
   (*Index through the event listing and get current value for each code*)
   (*The first element in the array is the array length*)
   FOR Index := 1 TO CCPSystem.EventList.Event[0] DO;
   
   	(*Extract the Structure, Tag and Property values from the code.  The code is in the format SSTTTPP*)
   	Code := CCPSystem.EventList.Event[Index];
   	DTOS (Code, sCode);
   
   		IF sCode.LEN = 7 THEN;
   			MID (sCode, 2, 1, sStructure);
   			MID (sCode, 3, 3, sTag);
   			MID (sCode, 2, 6, sProperty);
   		ELSIF sCode.LEN = 6 THEN;
   			MID (sCode, 1, 1, sStructure);
   			MID (sCode, 3, 2, sTag);
   			MID (sCode, 2, 5, sProperty);
   		ELSE;
   			(*Ignore if code length is not 6 or 7*)
   			DTOS (0, sStructure);
   		END_IF;
   		STOD (sStructure, Structure);
   		STOD (sTag, Tag);
   		STOD (sProperty, Property);
   
   	(* Tag:= 0; (*put in to handel error in congig files*)
   
   	Value := 0;
   
   (* Navigate through the event categories
   =========================================================================*)
   	(*Get the value based on the structure, tag and property*)
   	CASE	Structure OF
   		1: 	CASE	Property OF (*Analog Alarms*)
   			1:	IF AlarmAnalog[Tag].Override THEN Value := 1; ELSE Value := 0; END_IF;
   			2:	Value := AlarmAnalog[Tag].LOLO;
   			3:	Value := AlarmAnalog[Tag].LO;
   			4:	Value := AlarmAnalog[Tag].HI;
   			5:	Value := AlarmAnalog[Tag].HIHI;
   			6:	IF AlarmAnalog[Tag].LOLOAlarm THEN Value := 1; ELSE Value := 0; END_IF;
   			7:	IF AlarmAnalog[Tag].LOAlarm THEN Value := 1; ELSE Value := 0; END_IF;
   			8:	IF AlarmAnalog[Tag].HIAlarm THEN Value := 1; ELSE Value := 0; END_IF;
   			9:	IF AlarmAnalog[Tag].HIHIAlarm THEN Value := 1; ELSE Value := 0; END_IF;
   			END_CASE;
   		2: 	CASE	Property OF (*Deviation Alarms*)
   			1:	IF AlarmDeviation[Tag].Override THEN Value := 1; ELSE Value := 0; END_IF;
   			4:	Value := AlarmDeviation[Tag].HI;
   			5:	Value := AlarmDeviation[Tag].HIHI;
   			8:	IF AlarmDeviation[Tag].HIAlarm THEN Value := 1; ELSE Value := 0; END_IF;
   			9:	IF AlarmDeviation[Tag].HIHIAlarm THEN Value := 1; ELSE Value := 0; END_IF;
   			END_CASE;
   		3: 	CASE	Property OF (*Digital Alarms*)
   			1:	IF DigitalPoint[Tag].Override THEN Value := 1; ELSE Value := 0; END_IF;
   			6:	IF DigitalPoint[Tag].Alarm THEN Value := 1; ELSE Value := 0; END_IF;
   			7:	IF DigitalPoint[Tag].CurrentValue THEN Value := 1; ELSE Value := 0; END_IF;
   			END_CASE;
   		4: 	CASE	Property OF (*Analog Inputs*)
   			1:	Value := AnalogPoint[Tag].CurrentValue;
   			2:	Value := AnalogPoint[Tag].ScaledMin;
   			3:	Value := AnalogPoint[Tag].ScaledMax;
   			END_CASE;
   		5:	CASE	Property OF (*Control Loops*)
   			1:	IF ControlLoop[Tag].Manual THEN Value := 1; ELSE Value := 0; END_IF;
   			2:	IF ControlLoop[Tag].Auto1 THEN Value := 1; ELSE Value := 0; END_IF;
   			3:	IF ControlLoop[Tag].Auto2 THEN Value := 1; ELSE Value := 0; END_IF;
   			4:	IF ControlLoop[Tag].Auto3 THEN Value := 1; ELSE Value := 0; END_IF;
   			5:	IF ControlLoop[Tag].Auto4 THEN Value := 1; ELSE Value := 0; END_IF;
   			6:	Value := ControlLoop[Tag].SPManual;
   			7:	Value := ControlLoop[Tag].SPAuto1;
   			8:	Value := ControlLoop[Tag].SPAuto2;
   			9:	Value := ControlLoop[Tag].SPAuto3;
   			10:	Value := ControlLoop[Tag].SPAuto4;
   			11:	Value := ControlLoop[Tag].RampRate;
   			12:	Value := ControlLoop[Tag].Deadband;
   			13:	Value := ControlLoop[Tag].StableTime;
   			14:	Value := ControlLoop[Tag].KP[0];
   			15:	Value := ControlLoop[Tag].KI[0];
   			16:	Value := ControlLoop[Tag].KD[0];
   			17:	Value := ControlLoop[Tag].DB[0];
   			18:	Value := ControlLoop[Tag].KP[1];
   			19:	Value := ControlLoop[Tag].KI[1];
   			20:	Value := ControlLoop[Tag].KD[1];
   			21:	Value := ControlLoop[Tag].DB[1];
   			22:	Value := ControlLoop[Tag].KP[2];
   			23:	Value := ControlLoop[Tag].KI[2];
   			24:	Value := ControlLoop[Tag].KD[2];
   			25:	Value := ControlLoop[Tag].DB[2];
   			26:	IF ControlLoop[Tag].Stable THEN Value := 1; ELSE Value := 0; END_IF;
   			27:	IF ControlLoop[Tag].DBOK THEN Value := 1; ELSE Value := 0; END_IF;
   			28:	IF ControlLoop[Tag].RampStatus THEN Value := 1; ELSE Value := 0; END_IF;
   			END_CASE;
   		7:	CASE	Property OF (*Phase Control*)
   			1:	IF Phase[Tag].Run THEN Value := 1; ELSE Value := 0; END_IF;
   			2:	IF Phase[Tag].Stop THEN Value := 1; ELSE Value := 0; END_IF;
   			3:	IF Phase[Tag].Hold THEN Value := 1; ELSE Value := 0; END_IF;
   			4:	IF Phase[Tag].Pause THEN Value := 1; ELSE Value := 0; END_IF;
   			5:	IF Phase[Tag].Label = 0 THEN CCPSystem.EventList.Value[Index] := 0; END_IF; (*Ignore change to 0*)
   				Value := Phase[Tag].Label;
   			6:	IF Phase[Tag].JumpPLC THEN Value := 1; ELSE Value := 0; END_IF;
   			END_CASE;
   		8: 	CASE	Property OF (*Prompts*)
   			1:	IF Prompt[Tag].PromptOK THEN Value := 1; ELSE Value := 0; END_IF;
   			2:	IF Prompt[Tag].PromptYesNO THEN Value := 1; ELSE Value := 0; END_IF;
   			3:	IF Prompt[Tag].ResponseOK THEN Value := 1; ELSE Value := 0; END_IF;
   			4:	IF Prompt[Tag].ResponseYes THEN Value := 1; ELSE Value := 0; END_IF;
   			5:	IF Prompt[Tag].ResponseNo THEN Value := 1; ELSE Value := 0; END_IF;
   			END_CASE;
   		9: 	CASE	Property OF (*Pumps*)
   			1:	IF Drive[Tag].RunStatus THEN Value := 1; ELSE Value := 0; END_IF;
   			2:	IF Drive[Tag].Direction THEN Value := 1;ELSE Value := 0; END_IF;
   			3:	IF Drive[Tag].Mode THEN Value := 1; ELSE Value := 0; END_IF;
   			END_CASE;
   		11:	CASE	Property OF (*Timers*)
   			3:	IF Timers[Tag].Enable THEN Value := 1; ELSE Value := 0; END_IF;
   			4:	IF Timers[Tag].Reset THEN Value := 1; ELSE Value := 0; END_IF;
   			END_CASE;
   		13:	CASE	Property OF (*Valves*)
   			2:	Value := Valve[Tag].StatusWord;
   			3:	IF Valve[Tag].Mode THEN Value := 1; ELSE Value := 0; END_IF;
   			4:	IF Valve[Tag].Alarm THEN Value := 1; ELSE Value := 0; END_IF;
   			5:	Value := Valve[Tag].Status;
   			END_CASE;
   		14:	CASE	Property OF (*Agitator*)
   			1:	IF Mixer.Mode THEN Value := 1; ELSE Value := 0; END_IF;
   			2:	Value := Mixer.SPManual;
   			3:	Value := Mixer.SPAutoMin;
   			4:	Value := Mixer.SPAutoMax;
   			5:	Value := Mixer.LevelMin;
   			6:	Value := Mixer.LevelMax;
   			END_CASE;
   		15:	CASE	Property OF (*Misc.*)
   			1:	IF MiscBOOL[Tag] THEN Value := 1; ELSE Value := 0; END_IF;
   			2:	Value := MiscDINT[Tag];
   			3:	Value := MiscREAL[Tag];
   			END_CASE;
   		16:	CASE	Property OF (*Alarm Control*)
   			1:	IF AlarmControl.EnableAllOut THEN Value := 1; ELSE Value := 0; END_IF;
   			2:	IF AlarmControl.DisableAllOut THEN Value := 1; ELSE Value := 0; END_IF;
   			3:	IF AlarmControl.AckOutput THEN Value := 1; ELSE Value := 0; END_IF;
   			6:	IF AlarmControl.EnableAllAnaSigOut THEN Value := 1; ELSE Value := 0; END_IF;
   			7:	IF AlarmControl.DisableAllAnaSigOut THEN Value := 1; ELSE Value := 0; END_IF;
   			END_CASE;
   		17:	CASE	Property OF (*Miscellaneous*)
   			1:	IF SysControl.DefaultOut THEN Value := 1; ELSE Value := 0; END_IF;
   			2:	IF ChartMark.Out THEN Value := 1; ELSE Value := 0; END_IF;
   			3:	IF SysControl.AllAutoOut THEN Value := 1; ELSE Value := 0; END_IF;
   			4:	IF UserTotalizerManagement.LogUserOut THEN Value := 1; ELSE Value := 0; END_IF;
   			5:	IF UserTotalizerManagement.StartUser THEN Value := 1; ELSE Value := 0; END_IF;
   			6:	IF UserTotalizerManagement.ResetUserOut THEN Value := 1; ELSE Value := 0; END_IF;
   			7:	IF Tank.Feed_Bag_Tare THEN Value := 1; ELSE Value := 0; END_IF;
   			8:	IF Tank.Filtrate_Bag_Tare THEN Value := 1; ELSE Value := 0; END_IF;
   			9:	IF SysControl.UV_Auto_Zero_Cmd THEN Value := 1; ELSE Value := 0; END_IF;
   			11:	IF CCPSystem.DefaultOnComplete THEN Value := 1; ELSE Value := 0; END_IF;
   			12:	IF UserAlarm.NonCritical1 THEN Value := 1; ELSE Value := 0; END_IF;
   			13:	IF UserAlarm.Critical1 THEN Value := 1; ELSE Value := 0; END_IF;
   			14:	IF UserAlarm.NonCritical2 THEN Value := 1; ELSE Value := 0; END_IF;
   			15:	IF UserAlarm.Critical2 THEN Value := 1; ELSE Value := 0; END_IF;
   			16:	IF SRL001.CurrentValue THEN Value := 1; ELSE Value := 0; END_IF;
   			END_CASE;
   		18:	CASE	Property OF (*Criteria Flag*)
   			1:	IF CriteriaFlag.Flag1 THEN Value := 1; ELSE Value := 0; END_IF;
   			2:	IF CriteriaFlag.Flag2 THEN Value := 1; ELSE Value := 0; END_IF;
   			3:	IF CriteriaFlag.Flag3 THEN Value := 1; ELSE Value := 0; END_IF;
   			4:	IF CriteriaFlag.Flag4 THEN Value := 1; ELSE Value := 0; END_IF;
   			5:	IF CriteriaFlag.Flag5 THEN Value := 1; ELSE Value := 0; END_IF;
   			END_CASE;
   		19:	CASE	Property OF (*Concentration*)
   			1:	IF FQ_Conc.Enable THEN Value := 1; ELSE Value := 0; END_IF;
   			2:	IF FQ_Conc.Reset THEN Value := 1; ELSE Value := 0; END_IF;
   			3:	IF Concentration.LogConcOut THEN Value := 1; ELSE Value := 0; END_IF;
   			4:	Value := Concentration.Conc_Init ;
   			5:	Value := Concentration.Conc_Final ;
   			6:	Value := Concentration.Conc_Final_Volume ;
   			7:	Value := DerivedData.HOLDUP ;
   			10: IF Concentration.Final_Conc_Volume_Reached THEN Value := 1; ELSE Value := 0; END_IF;
   			11: IF Concentration.Final_Conc_Protein_Reached THEN Value := 1; ELSE Value := 0; END_IF;
   			END_CASE;
   		20:	CASE	Property OF (*Diafiltration*)
   			1:	IF FQ_Diaf.Enable THEN Value := 1; ELSE Value := 0; END_IF;
   			2:	IF FQ_Diaf.Reset THEN Value := 1; ELSE Value := 0; END_IF;
   			3:	IF Diafiltration.LogDiafOut THEN Value := 1; ELSE Value := 0; END_IF;
   			4:	IF Diafiltration.Snap THEN Value := 1; ELSE Value := 0; END_IF;
   			5:	Value := Diafiltration.Diaf_Init ;
   			6:	Value := Diafiltration.Diaf_Final_Volume ;
   			10: IF Diafiltration.Final_Diaf_Volum_Reached THEN Value := 1; ELSE Value := 0; END_IF;
   			END_CASE;
   		21:	CASE	Property OF (*Membrane Data*)
   			1:	Value := Membrane_Data.Area ;
   			2:	Value := Membrane_Data.Density ;
   			END_CASE;
   		23:	CASE	Property OF (*PCV Control*)
   			1:	IF PCV001_Control.FullOpen THEN Value := 1; ELSE Value := 0; END_IF;
   			2:	IF PCV001_Control.FullClose THEN Value := 1; ELSE Value := 0; END_IF;
   			3:	IF PCV101_Control.FullOpen THEN Value := 1; ELSE Value := 0; END_IF;
   			4:	IF PCV101_Control.FullClose THEN Value := 1; ELSE Value := 0; END_IF;
   			END_CASE;
   		24:	CASE	Property OF (*Event value.*)
   			1:	Value := LogVal.Value[Tag];
   			END_CASE;
   		25: CASE	Property OF (*Flow Paths*)
   			1:	IF FlowPath[Tag].Status THEN Value := 1; ELSE Value := 0; END_IF;
   			2:	IF FlowPathControl.FlushMode_Enabled THEN Value := 1; ELSE Value := 0; END_IF;
   			3:	IF FlowPathControl.DrainMode_Enabled THEN Value := 1; ELSE Value := 0; END_IF;
   			END_CASE;
   		26: CASE	Property OF (*Clamshell*)
   			1:	IF Y500A THEN Value := 1; ELSE Value := 0; END_IF;
   			2:	IF Y500B THEN Value := 1; ELSE Value := 0; END_IF;
   			3:	IF Y501A THEN Value := 1; ELSE Value := 0; END_IF;
   			4:	IF Y501B THEN Value := 1; ELSE Value := 0; END_IF;
   			5:	IF Y502A THEN Value := 1; ELSE Value := 0; END_IF;
   			6:	IF Y502B THEN Value := 1; ELSE Value := 0; END_IF;
   			7:	IF Y503A THEN Value := 1; ELSE Value := 0; END_IF;
   			8:	IF Y503B THEN Value := 1; ELSE Value := 0; END_IF;
   			11:  IF ThisSystem.MoldType = 123 THEN Value := 1; ELSE Value := 0; END_IF;
   			12:  IF ThisSystem.MoldType = 124 THEN Value := 1; ELSE Value := 0; END_IF;
   			21:  IF ThisSystem.PreviousValue = 123 THEN Value := 1; ELSE Value := 0; END_IF;
   			22:  IF ThisSystem.PreviousValue = 124 THEN Value := 1; ELSE Value := 0; END_IF;
   			END_CASE;
   		30:	CASE	Property OF (*DCS Actions Events*)
   			0:	Value := DCS.ActionsParameters.Feed_Pump_Speed_Setpoint[Tag];
   			1:	Value := DCS.ActionsParameters.Feed_Pump_Flow_Setpoint[Tag];
   			2:	Value := DCS.ActionsParameters.Feed_Pump_DP_Setpoint[Tag];
   			3:	Value := DCS.ActionsParameters.Level_Pump_Speed_Setpoint[Tag];
   			4:	Value := DCS.ActionsParameters.Level_Pump_Level_Setpoint[Tag];
   			6:	Value := DCS.ActionsParameters.PCV001_Retentate_Position_Setpoint[Tag];
   			7:	Value := DCS.ActionsParameters.PCV001_Retentate_Pressure_Setpoint[Tag];
   			8:	Value := DCS.ActionsParameters.PCV001_Retentate_TMP_Setpoint[Tag];
   			9:	Value := DCS.ActionsParameters.PCV101_Filtrate_Position_Setpoint[Tag];
   			10:	Value := DCS.ActionsParameters.PCV101_Filtrate_Flow_Setpoint[Tag];
   			11:	Value := DCS.ActionsParameters.PCV101_Filtrate_TMP_Setpoint[Tag];
   			12:	Value := DCS.ActionsParameters.Mixer_Speed_Setpoint[Tag];
   			13:	Value := DCS.ActionsParameters.Mixer_Auto_Min_Setpoint[Tag];
   			14:	Value := DCS.ActionsParameters.Mixer_Auto_Max_Setpoint[Tag];
   			15:	Value := DCS.ActionsParameters.Init_Protein_Conc[Tag];
   			16:	Value := DCS.ActionsParameters.Final_Protein_Conc[Tag];
   			17:	Value := DCS.ActionsParameters.Final_Protein_Volume[Tag];
   			18:	Value := DCS.ActionsParameters.Holdup_Volume[Tag];
   			19:	Value := DCS.ActionsParameters.Init_Diaf_Volume[Tag];
   			20:	Value := DCS.ActionsParameters.Final_Diaf_Volume[Tag];
   			21:	Value := DCS.ActionsParameters.Membrane_Area[Tag];
   			22:	Value := DCS.ActionsParameters.Membrane_Density[Tag];
   			END_CASE;
   	31: CASE	Property OF (*DCS Criteria*)
   			1:	IF DCS.Criteria.Criteria_1 THEN Value := 1; ELSE Value := 0; END_IF;
   			2:	IF DCS.Criteria.Criteria_2 THEN Value := 1; ELSE Value := 0; END_IF;
   			END_CASE;
   	(*Missing else statement accepted for the purpose of proper integration with CCPRuntime.exe*)
   	END_CASE;
   
   (* Log Pre-run values
   =========================================================================*)
   	(*Record value for Pre-Run Log if flag is set*)
   	IF PreRunLog THEN;
   		CCPSystem.EventList.PreRunValue[Index] := Value;
   	END_IF;
   
   
   (* Build event contents
   =========================================================================*)
   	(*Check for change in value*)
   	IF CCPSystem.EventList.Value[Index] <> Value THEN;
   		(*Increment pointer*)
   		Pointer := Pointer + 1;
   		(*Roll over pointer if equal to max*)
   		IF Pointer = 251 THEN Pointer := 1; END_IF;
   
   		(*Concatenate the action code to the date/time and add comma*)
   		DTOS (Code, sTemp);
   		CONCAT(sDateTime, sTemp, sBufferEvents);
   		CONCAT(sBufferEvents, sComma, sBufferEvents);
   
   		(*Concatenate the new value and add comma*)
   		RTOS (Value, sTemp);
   		CONCAT (sBufferEvents, sTemp, sBufferEvents);
   		CONCAT (sBufferEvents, sComma, sBufferEvents);
   
   		(*Concatenate the old value and store in the buffer*)
   		RTOS(CCPSystem.EventList.Value[Index], sTemp);
   		CONCAT(sBufferEvents, sTemp, CCPSystem.BufferEvents[Pointer]);
   
   		(*Clear the unused characters for null termination*)
   		TempEvents := CCPSystem.BufferEvents[Pointer].LEN;
   		WHILE TempEvents < 50 DO;
   			CCPSystem.BufferEvents[Pointer].DATA[TempEvents] := 0;
   			TempEvents := TempEvents + 1;
   		END_WHILE;
   
   		(*Save the new value for subsequent comparison*)
   		CCPSystem.EventList.Value[Index] := Value;
   	END_IF;
   END_FOR;
   
   (* Reset flag and pointer
   =========================================================================*)
   (*Clear the pre-run log flag*)
   PreRunLog := 0;
   
   (*Update the buffer pointer value after processing all events*)
   DTOS (Pointer, CCPSystem.BufferEvents[0]);
   
END_ROUTINE

ROUTINE BufferSteps   (* structured text *)
// Step Log Buffer Routine
   (* =======================================================================
   	Buffer Steps : This routine updates the step buffer when a step is executed
   
   	List of treatments
   		- Get current action code
   		- Compute the step value for the step buffer
   
   -----------------------------------------------------------------------------------------------------------------------------------------------------
   	History
   		2019-AUG-13 - ACTEMIUM - B. Roch - Initial version for Candidate Release 3.00.00.00.a
   		2023-FEB-07 - Davidson - Ch.Arbogast - Modifications for Candidate Release 3.02.00.00.a
   					- Limit LastStep to 0 minimum after "LastStep := PendingStep - 1;"
   							add " IF LastStep < 0 THEN;	LastStep := 0; END_IF;"
   =========================================================================*)
   
   
   (* Get the current pointer value and increment
   =========================================================================*)
   STOD (CCPSystem.BufferSteps[0], Pointer);
   Pointer := Pointer + 1;
   (*Roll over pointer if equal to max*)
   IF Pointer = 251 THEN Pointer := 1; END_IF;
   DTOS (Pointer, CCPSystem.BufferSteps[0]);
   
   (* Compute the step value for the step buffer
   =========================================================================*)
   (*If the pending step number is the same as the last step number (named action list) then add 10000 to the buffer value*)
   LastStep := PendingStep - 1;
   IF LastStep < 0 THEN;
   	LastStep := 0;
   END_IF;
   IF Operation[PhaseNumber,PendingStep].Step = Operation[PhaseNumber,LastStep].Step THEN;
   	BufferStep := PhaseNumber * 1000 + (Operation[PhaseNumber,PendingStep].Step) + 10000;
   ELSE;
   	BufferStep := PhaseNumber * 1000 + (Operation[PhaseNumber,PendingStep].Step);
   END_IF;
   
   (*Convert the step value to a string and concatenate with the date/time*)
   DTOS (BufferStep, sTemp);
   CONCAT (sDateTime, sTemp, CCPSystem.BufferSteps[Pointer]);
   
   (*Clear the unused characters for null termination*)
   TempSteps := CCPSystem.BufferSteps[Pointer].LEN;
   WHILE TempSteps < 26 DO;
   	CCPSystem.BufferSteps[Pointer].DATA[TempSteps] := 0;
   	TempSteps := TempSteps + 1;
   END_WHILE;
END_ROUTINE

ROUTINE Clear   (* structured text *)
// Clear Operation Table
   (* =======================================================================
   	Clear : This routine loops through the entire operation array and clears
   			the step numbers, set Criteria1Value, Criteria2Value, ActionValue
   			to -999999.99 and sets all other values to -999.
   			This is executed at the start of each download.
   
   	List of treatments
   		- Initialize phase clear number
   		- Reset Operation data
   		- Reset Prompt messages
   		- In case of procedure RunAuto flag is set
   
   -----------------------------------------------------------------------------------------------------------------------------------------------------
   	History
   		2019-AUG-13 - ACTEMIUM - B. Roch - Initial version for Candidate Release 3.00.00.00.a
   		2019-SEP-09 - ACTEMIUM - Q. Spindler - Modifications for Candidate Release 3.00.00.00.c
   					- Change Error check for Criterias and Action Value to -999999.99
   =========================================================================*)
   
   
   (* Initialize phase clear number
   =========================================================================*)
   (*One-Shot to set phase clear number to zero*)
   IF NOT PhaseClear THEN;
   	PhaseClearNumber := 0;
   	PhaseClear := 1;
   END_IF;
   
   (* Reset Operation data
   =========================================================================*)
   (*Step FOR-NEXT loop*)
   FOR PendingStep := 1 TO 250 DO;
   	Operation [PhaseClearNumber, PendingStep].Step := 0;
   	Operation [PhaseClearNumber, PendingStep].Criteria1 := -999;
   	Operation [PhaseClearNumber, PendingStep].Criteria1Operator := -999;
   	Operation [PhaseClearNumber, PendingStep].Boolean := -999;
   	Operation [PhaseClearNumber, PendingStep].Criteria2 := -999;
   	Operation [PhaseClearNumber, PendingStep].Criteria2Operator := -999;
   	Operation [PhaseClearNumber, PendingStep].Action := -999;
   	Operation [PhaseClearNumber, PendingStep].Label := -999;
   	Operation [PhaseClearNumber, PendingStep].Criteria1Value := -999999.99;
   	Operation [PhaseClearNumber, PendingStep].Criteria2Value := -999999.99;
   	Operation [PhaseClearNumber, PendingStep].ActionValue := -999999.99;
   END_FOR;
   
   PhaseClearNumber := PhaseClearNumber + 1;
   
   (* Reset Prompt messages
   =========================================================================*)
   IF PhaseClearNumber = 6 THEN;
   	(*Clear step buffer*)
   	CCPSystem.BufferSteps[0].LEN := 0;
   	(*State 11 ready for download*)
   	CCPSystem.State := 11;
   
   	Prompt0.PromptOK := 0;
   	Prompt0.PromptYesNO := 0;
   	Prompt1.PromptOK := 0;
   	Prompt1.PromptYesNO := 0;
   	Prompt2.PromptOK := 0;
   	Prompt2.PromptYesNO := 0;
   	Prompt3.PromptOK := 0;
   	Prompt3.PromptYesNO := 0;
   	Prompt4.PromptOK := 0;
   	Prompt4.PromptYesNO := 0;
   	Prompt5.PromptOK := 0;
   	Prompt5.PromptYesNO := 0;
   
   (* In case of procedure RunAuto flag is set
   =========================================================================*)
   	(*If part of a procedure then set the auto run flag so the operation will start when download is completed*)
   	IF CCPSystem.Procedure THEN;
   		CCPSystem.RunAuto := 1;
   	ELSE;
   		CCPSystem.RunAuto := 0;
   	END_IF;
   
   	PhaseClear := 0;
   
   END_IF;
   
END_ROUTINE

ROUTINE Complete   (* ladder *)
// Operation Complete Routine
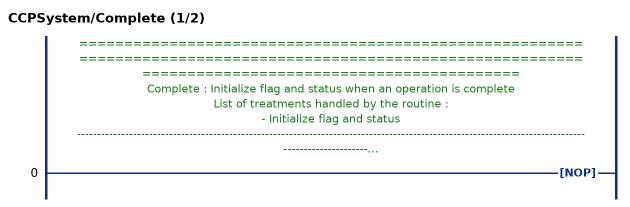
   // ==========================================================================================================================================================
   //                                                                                                Complete : Initialize flag and status when an operation is complete
   //                                                     List of treatments handled by the routine :
   //                                                          - Initialize flag and status
   //                                                     -----------------------------------------------------------------------------------------------------------------------------------------------------
   //                                                     History
   //                                                          2019-AUG-13 - Actemium - B. Roch - Initial version for Candidate Release 3.00.00.00.a
   // 		2022-FEB-02 - Davidson - Ch.Arbogast - Modifications for Candidate Release 3.02.00.00.a
   // 				- Add unlatch of CCPSystem.Procedure when procedure is aborted
   // ========================================================================================================================================================
   0: NOP();
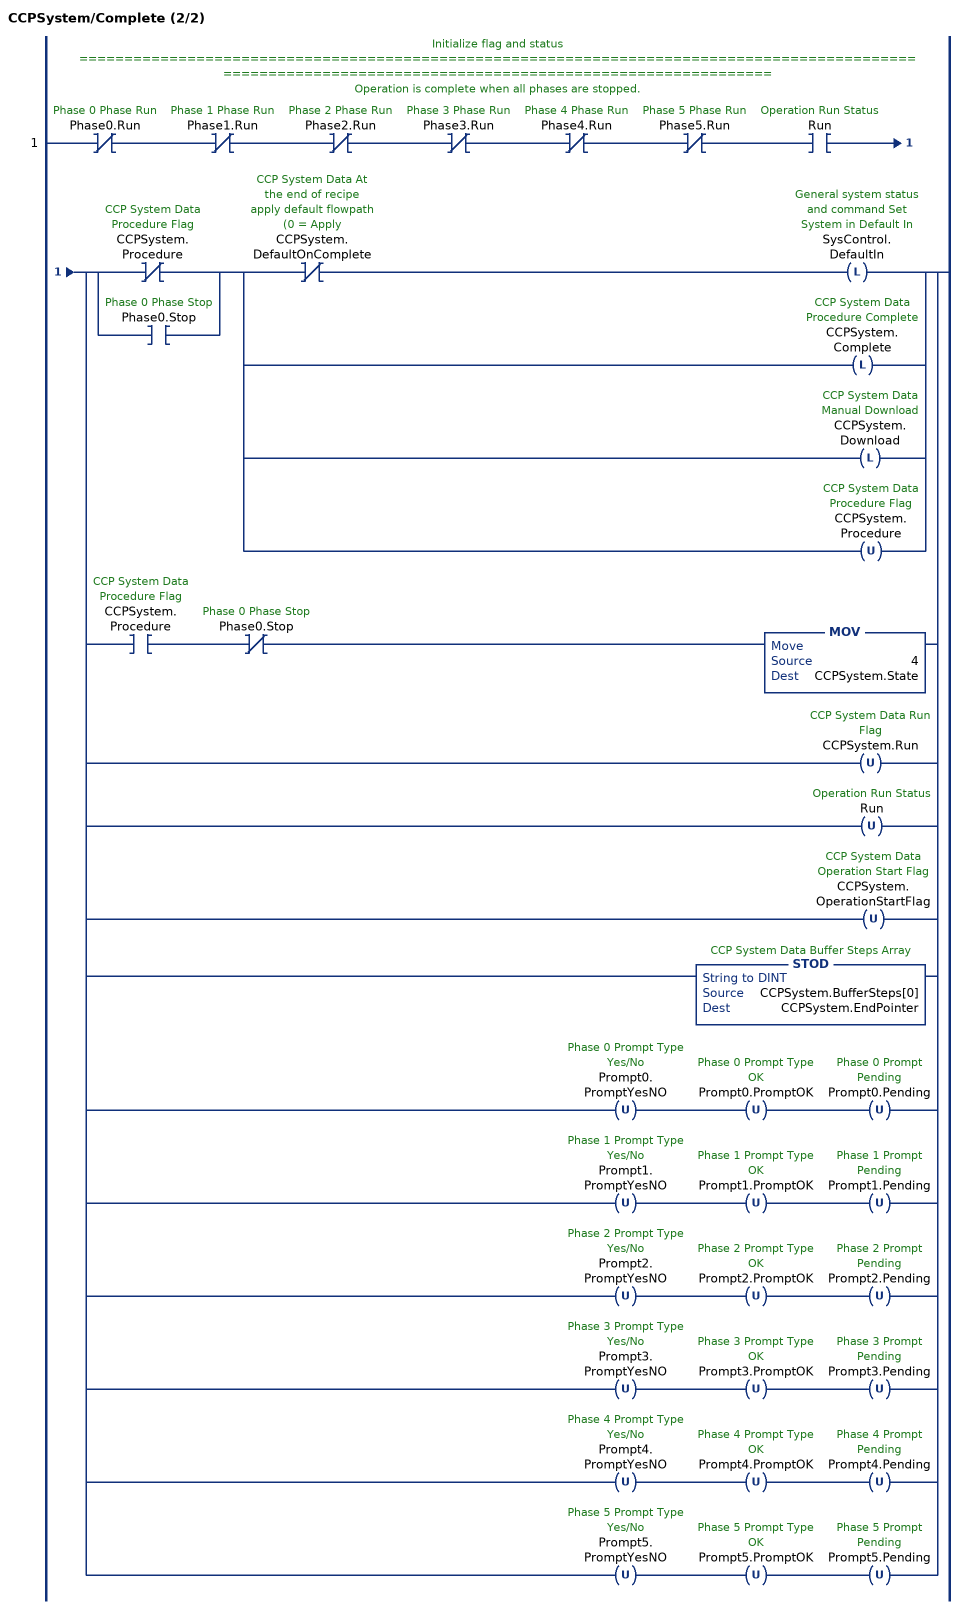
   // Initialize flag and status
   // ==========================================================================================================================================================
   // Operation is complete when all phases are stopped.
   1: XIO(Phase0.Run)XIO(Phase1.Run)XIO(Phase2.Run)XIO(Phase3.Run)XIO(Phase4.Run)XIO(Phase5.Run)XIC(Run)[[XIO(CCPSystem.Procedure) ,XIC(Phase0.Stop) ] [XIO(CCPSystem.DefaultOnComplete) OTL(SysControl.DefaultIn) ,OTL(CCPSystem.Complete) ,OTL(CCPSystem.Download) ,OTU(CCPSystem.Procedure) ] ,XIC(CCPSystem.Procedure) XIO(Phase0.Stop) MOV(4,CCPSystem.State) ,OTU(CCPSystem.Run) ,OTU(Run) ,OTU(CCPSystem.OperationStartFlag) ,STOD(CCPSystem.BufferSteps[0],CCPSystem.EndPointer) ,OTU(Prompt0.PromptYesNO) OTU(Prompt0.PromptOK) OTU(Prompt0.Pending) ,OTU(Prompt1.PromptYesNO) OTU(Prompt1.PromptOK) OTU(Prompt1.Pending) ,OTU(Prompt2.PromptYesNO) OTU(Prompt2.PromptOK) OTU(Prompt2.Pending) ,OTU(Prompt3.PromptYesNO) OTU(Prompt3.PromptOK) OTU(Prompt3.Pending) ,OTU(Prompt4.PromptYesNO) OTU(Prompt4.PromptOK) OTU(Prompt4.Pending) ,OTU(Prompt5.PromptYesNO) OTU(Prompt5.PromptOK) OTU(Prompt5.Pending) ];
END_ROUTINE

ROUTINE Criteria1   (* structured text *)
// Criteria 1 Routine
   (* =======================================================================
   	Criteria1 : Get the current criteria 1 code and verify if criteria met based on information extraction.
   				Update the criteria 1 bool and real value and the criteria type.
   
   	List of treatments
   		- Initialize Phase step number
   		- Extract informations based on criteria 1 code
   		- Navigate through the criteria categories and set Criteria bool and real value
   
   -----------------------------------------------------------------------------------------------------------------------------------------------------
   	History
   		2019-AUG-13 - ACTEMIUM - B. Roch - Initial version for Candidate Release 3.00.00.00.a
   		2020-SEP-21 - Merck - Q. Spindler - Modifications for Candidate Release 3.00.00.01.a
   			- Remove Criteria1Type := 1 for VCF, CB, and Diaf_Volume (As they are Real Criteria)
   		2021-MAY-03 - DAVIDSON- Ch. ARBOGAST - Modifications for Candidate Release 3.01.00.00.a
    			- on case 11,line 1:,add test  "IF Timers[Criteria1Tag].Reset THEN Criteria1RealValue := 0;"
   		2023-FEB-14 - Davidson - Ch.Arbogast - Modifications for Candidate Release 3.02.00.00.a
   			- add Case 30: DCS criteria
   =========================================================================*)
   
   (* Initialize Phase step number
   =========================================================================*)
   (*If error check, pending step number is set by error check loop*)
   IF NOT ErrorCheck THEN;
   	PendingStep := Phase[PhaseNumber].ActualStep;
   	Phase[PhaseNumber].PendingStep := Operation[PhaseNumber,PendingStep].Step;
   	NextStep := PendingStep + 1;
   	IF PendingStep < 250 AND Operation[PhaseNumber,NextStep].Step <> 0 THEN;
   		Phase[PhaseNumber].NextStep := Operation[PhaseNumber,NextStep].Step;
   	ELSE;
   		Phase[PhaseNumber].NextStep := 0;
   	END_IF;
   END_IF;
   
   (* Extract informations based on criteria 1 code
   =========================================================================*)
   Criteria1Code := Operation[PhaseNumber,PendingStep].Criteria1;
   Criteria1Operator := Operation[PhaseNumber,PendingStep].Criteria1Operator;
   Criteria1Value := Operation[PhaseNumber,PendingStep].Criteria1Value;
   Boolean := Operation[PhaseNumber,PendingStep].Boolean;
   Criteria1Type := 0;
   
   (*Extract the Structure, Tag and Property values from the criteria code.  The criteria code is
   in the format SSTTTPP*)
   
   IF Criteria1Code <> 0 THEN;
   	DTOS (Criteria1Code, sCriteria1);
   	IF sCriteria1.LEN = 7 THEN;
   		MID (sCriteria1, 2, 1, sCriteria1Structure);
   		MID (sCriteria1, 3, 3, sCriteria1Tag);
   		MID (sCriteria1, 2, 6, sCriteria1Property);
   	ELSIF sCriteria1.LEN = 6 THEN;
   		MID (sCriteria1, 1, 1, sCriteria1Structure);
   		MID (sCriteria1, 3, 2, sCriteria1Tag);
   		MID (sCriteria1, 2, 5, sCriteria1Property);
   	ELSE;
   		CCPSystem.Error := 2;
   	END_IF;
   	STOD (sCriteria1Structure, Criteria1Structure);
   	STOD (sCriteria1Tag, Criteria1Tag);
   	STOD (sCriteria1Property, Criteria1Property);
   ELSE;
   	Criteria1Structure := 0;
   END_IF;
   
   (* Navigate through the criteria categories and set Criteria bool and real value
   =========================================================================*)
   CASE	Criteria1Structure OF
   	0:	; (*No Criteria*)
   	3:	CASE	Criteria1Property OF (*Digital Points*)
   			1:	Criteria1BoolValue := DigitalPoint[Criteria1Tag].CurrentValue;
   				Criteria1Type := 1;
   			2:	Criteria1BoolValue := DigitalPoint[Criteria1Tag].Alarm;
   				Criteria1Type := 1;
   			3:	Criteria1BoolValue := DigitalPoint[Criteria1Tag].SoftInput;
   				Criteria1Type := 1;
   		ELSE 	CCPSystem.Error := 2;
   		END_CASE;
   	4: 	CASE	Criteria1Property OF (*Analog Inputs*)
   			1:	Criteria1RealValue := AnalogPoint[Criteria1Tag].CurrentValue;
   		ELSE 	CCPSystem.Error := 2;
   		END_CASE;
   	5:	CASE	Criteria1Property OF (*Control Loops*)
   			18:	Criteria1BoolValue := ControlLoop[Criteria1Tag].Stable;
   				Criteria1Type := 1;
   			19:	Criteria1BoolValue := ControlLoop[Criteria1Tag].DBOK;
   				Criteria1Type := 1;
   			20:	Criteria1BoolValue := ControlLoop[Criteria1Tag].RampStatus;
   				Criteria1Type := 1;
   		ELSE 	CCPSystem.Error := 2;
   		END_CASE;
   	7:	CASE	Criteria1Property OF (*Phase Control*)
   			1:	Criteria1BoolValue := Phase[Criteria1Tag].Run;
   				Criteria1Type := 1;
   			3:	Criteria1BoolValue := Phase[Criteria1Tag].Hold;
   				Criteria1Type := 1;
   			4:	Criteria1BoolValue := Phase[Criteria1Tag].Pause;
   		ELSE 	CCPSystem.Error := 2;
   		END_CASE;
   	8: 	CASE	Criteria1Property OF (*Prompts*)
   			3:	Criteria1BoolValue := Prompt[PhaseNumber].ResponseOK;
   				Criteria1Type := 1;
   			4:	Criteria1BoolValue := Prompt[PhaseNumber].ResponseYes;
   				Criteria1Type := 1;
   			5:	Criteria1BoolValue := Prompt[PhaseNumber].ResponseNo;
   				Criteria1Type := 1;
   		ELSE 	CCPSystem.Error := 2;
   		END_CASE;
   	9: 	CASE	Criteria1Property OF (*Pumps*)
   			2:	Criteria1BoolValue := Drive[Criteria1Tag].RunStatus;
   				Criteria1Type := 1;
   		ELSE 	CCPSystem.Error := 2;
   		END_CASE;
   	11:	CASE	Criteria1Property OF (*Timers*)
   			1:  IF Timers[Criteria1Tag].Reset THEN Criteria1RealValue := 0;
                   ELSE Criteria1RealValue := Timers[Criteria1Tag].TotalSeconds; (*Total Time*) END_IF;
   			2:	Criteria1Tag := Criteria1Tag + PhaseNumber; (*Add phase number to address correct step timer*)
   				Criteria1RealValue := Timers[Criteria1Tag].TotalSeconds; (*Step Time*)
   		ELSE 	CCPSystem.Error := 2;
   		END_CASE;
   	12:	CASE	Criteria1Property OF (*Totalizers*)
   			1:	Criteria1RealValue := PhaseTotalizer[Criteria1Tag].Phase;
   			2:	Criteria1Tag := Criteria1Tag + PhaseNumber; (*Add phase number to address correct step totalizer*)
   				Criteria1RealValue := PhaseTotalizer[Criteria1Tag].Step;
   			3:	Criteria1RealValue := PhaseTotalizer[Criteria1Tag].Pause;
   			4:	Criteria1RealValue := PhaseTotalizer[Criteria1Tag].User;
   			5:	Criteria1RealValue := PhaseTotalizer[Criteria1Tag].Procedure;
   			8:	Criteria1RealValue := Totalizer[Criteria1Tag].Total;
   		ELSE 	CCPSystem.Error := 2;
   		END_CASE;
   	13:	CASE	Criteria1Property OF (*Valves*)
   			2:	Criteria1RealValue := Valve[Criteria1Tag].StatusWord;
   		ELSE 	CCPSystem.Error := 2;
   		END_CASE;
   	15:	CASE	Criteria1Property OF (*Misc.*)
   			1:	Criteria1BoolValue := MiscBOOL[Criteria1Tag];
   				Criteria1Type := 1;
   			2:	Criteria1RealValue := MiscDINT[Criteria1Tag];
   			3:	Criteria1RealValue := MiscREAL[Criteria1Tag];
   		ELSE 	CCPSystem.Error := 2;
   		END_CASE;
   	17:	CASE	Criteria1Property OF (*Miscellaneous*)
   			11:	Criteria1BoolValue := CCPSystem.DefaultOnComplete ;
   				Criteria1Type := 1;
   		ELSE 	CCPSystem.Error := 2;
   		END_CASE;
   	18:	CASE	Criteria1Property OF (*Criteria Flag*)
   			1:	Criteria1BoolValue := CriteriaFlag.Flag1 ;
   				Criteria1Type := 1;
   			2:	Criteria1BoolValue := CriteriaFlag.Flag2 ;
   				Criteria1Type := 1;
   			3:	Criteria1BoolValue := CriteriaFlag.Flag3 ;
   				Criteria1Type := 1;
   			4:	Criteria1BoolValue := CriteriaFlag.Flag4 ;
   				Criteria1Type := 1;
   			5:	Criteria1BoolValue := CriteriaFlag.Flag5 ;
   				Criteria1Type := 1;
   		ELSE 	CCPSystem.Error := 2;
   		END_CASE;
   	19:	CASE	Criteria1Property OF (*Concentration*)
   			1:	Criteria1RealValue := Concentration.VCF;
   			2:	Criteria1RealValue := Concentration.CB;
   			3:	Criteria1BoolValue := Concentration.Final_Conc_Volume_Reached ;
   				Criteria1Type := 1;
   			4:	Criteria1BoolValue := Concentration.Final_Conc_Protein_Reached ;
   				Criteria1Type := 1;
   		ELSE 	CCPSystem.Error := 2;
   		END_CASE;
   	20:	CASE	Criteria1Property OF (*Diafiltration*)
   			1:	Criteria1RealValue := Diafiltration.Diaf_Volume;
   			2:	Criteria1BoolValue := Diafiltration.Final_Diaf_Volum_Reached ;
   				Criteria1Type := 1;
   		ELSE 	CCPSystem.Error := 2;
   		END_CASE;
   	25: CASE	Criteria1Property OF (*Flow Paths*)
   			2:	Criteria1BoolValue := FlowPath[Criteria1Tag].Status;
   				Criteria1Type := 1;
   		ELSE 	CCPSystem.Error := 2;
   		END_CASE;
   	30: CASE	Criteria1Tag OF (*DCS*)
   			0:	Criteria1BoolValue := DCS.Criteria.Criteria_1;
   				Criteria1Type := 1;
   			1:	Criteria1BoolValue := DCS.Criteria.Criteria_2;
   				Criteria1Type := 1;
   		ELSE 	CCPSystem.Error := 2;
   		END_CASE;
   ELSE	CCPSystem.Error := 2;
   END_CASE;
   
END_ROUTINE

ROUTINE Criteria2   (* structured text *)
// Criteria 2 Routine
   (* =======================================================================
   	Criteria2 : Get the current criteria 2 code and verify if criteria met based on information extraction.
   				Update the criteria 2 bool and real value and the criteria type.
   
   	List of treatments
   		- Initialize Phase step number
   		- Extract informations based on criteria 2 code
   		- Navigate through the criteria categories and set Criteria bool and real value
   
   -----------------------------------------------------------------------------------------------------------------------------------------------------
   	History
   		2019-AUG-13 - ACTEMIUM - B. Roch - Initial version for Candidate Release 3.00.00.00.a
   		2020-SEP-21 - Merck - Q. Spindler - Modifications for Candidate Release 3.00.00.01.a
   			- Remove Criteria2Type := 1 for VCF, CB, and Diaf_Volume (As they are Real Criteria)
   		2021-MAY-03 - DAVIDSON- Ch. ARBOGAST - Modifications for Candidate Release 3.01.00.00.a
    			- on case 11,line 1:,add test  "IF Timers[Criteria1Tag].Reset THEN Criteria1RealValue := 0;"
   		2023-FEB-14 - Davidson - Ch.Arbogast - Modifications for Candidate Release 3.02.00.00.a
   			- add Case 30: DCS criteria
   =========================================================================*)
   
   (* Extract informations based on criteria 2 code
   =========================================================================*)
   Criteria2Code := Operation[PhaseNumber,PendingStep].Criteria2;
   Criteria2Operator := Operation[PhaseNumber,PendingStep].Criteria2Operator;
   Criteria2Value := Operation[PhaseNumber,PendingStep].Criteria2Value;
   Criteria2Type := 0;
   
   IF Criteria2Code <> 0 THEN;
   	DTOS (Criteria2Code, sCriteria2);
   	IF sCriteria2.LEN = 7 THEN;
   		MID (sCriteria2, 2, 1, sCriteria2Structure);
   		MID (sCriteria2, 3, 3, sCriteria2Tag);
   		MID (sCriteria2, 2, 6, sCriteria2Property);
   	ELSIF sCriteria2.LEN = 6 THEN;
   		MID (sCriteria2, 1, 1, sCriteria2Structure);
   		MID (sCriteria2, 3, 2, sCriteria2Tag);
   		MID (sCriteria2, 2, 5, sCriteria2Property);
   	ELSE;
   		CCPSystem.Error := 5;
   	END_IF;
   	STOD (sCriteria2Structure, Criteria2Structure);
   	STOD (sCriteria2Tag, Criteria2Tag);
   	STOD (sCriteria2Property, Criteria2Property);
   ELSE;
   	Criteria2Structure := 0;
   END_IF;
   
   (* Navigate through the criteria categories and set Criteria bool and real value
   =========================================================================*)
   CASE	Criteria2Structure OF
   	0:	; (*No Criteria*)
   	3:	CASE	Criteria2Property OF (*Digital Points*)
   			1:	Criteria2BoolValue := DigitalPoint[Criteria2Tag].CurrentValue;
   				Criteria2Type := 1;
   			2:	Criteria2BoolValue := DigitalPoint[Criteria2Tag].Alarm;
   				Criteria2Type := 1;
   			3:	Criteria2BoolValue := DigitalPoint[Criteria2Tag].SoftInput;
   				Criteria2Type := 1;
   		ELSE 	CCPSystem.Error := 2;
   		END_CASE;
   	4: 	CASE	Criteria2Property OF (*Analog Inputs*)
   			1:	Criteria2RealValue := AnalogPoint[Criteria2Tag].CurrentValue;
   		ELSE 	CCPSystem.Error := 5;
   		END_CASE;
   	5:	CASE	Criteria2Property OF (*Control Loops*)
   			18:	Criteria2BoolValue := ControlLoop[Criteria2Tag].Stable;
   				Criteria2Type := 1;
   			19:	Criteria2BoolValue := ControlLoop[Criteria2Tag].DBOK;
   				Criteria2Type := 1;
   			20:	Criteria2BoolValue := ControlLoop[Criteria2Tag].RampStatus;
   				Criteria2Type := 1;
   		ELSE 	CCPSystem.Error := 5;
   		END_CASE;
   	7:	CASE	Criteria2Property OF (*Phase Control*)
   			1:	Criteria2BoolValue := Phase[Criteria2Tag].Run;
   				Criteria2Type := 1;
   			3:	Criteria2BoolValue := Phase[Criteria2Tag].Hold;
   				Criteria2Type := 1;
   			4:	Criteria2BoolValue := Phase[Criteria2Tag].Pause;
   			6:	Criteria2Tag := Criteria2Tag + PhaseNumber;
   				Criteria2RealValue := Phase[Criteria2Tag].Crit1MetTime;
   		ELSE 	CCPSystem.Error := 5;
   		END_CASE;
   	8: 	CASE	Criteria2Property OF (*Prompts*)
   			3:	Criteria2BoolValue := Prompt[PhaseNumber].ResponseOK;
   				Criteria2Type := 1;
   			4:	Criteria2BoolValue := Prompt[PhaseNumber].ResponseYes;
   				Criteria2Type := 1;
   			5:	Criteria2BoolValue := Prompt[PhaseNumber].ResponseNo;
   				Criteria2Type := 1;
   		ELSE 	CCPSystem.Error := 5;
   		END_CASE;
   	9: 	CASE	Criteria2Property OF (*Pumps*)
   			2:	Criteria2BoolValue := Drive[Criteria2Tag].RunStatus;
   				Criteria2Type := 1;
   		ELSE 	CCPSystem.Error := 5;
   		END_CASE;
   	11:	CASE	Criteria2Property OF (*Timers*)
   			1:  IF Timers[Criteria1Tag].Reset THEN Criteria1RealValue := 0;
                   ELSE Criteria1RealValue := Timers[Criteria1Tag].TotalSeconds; (*Total Time*) END_IF;
   			2:	Criteria2Tag := Criteria2Tag + PhaseNumber; (*Add phase number to address correct step timer*)
   				Criteria2RealValue := Timers[Criteria2Tag].TotalSeconds; (*Step Time*)
   		ELSE 	CCPSystem.Error := 5;
   		END_CASE;
   	12:	CASE	Criteria2Property OF (*Totalizers*)
   			1:	Criteria2RealValue := PhaseTotalizer[Criteria2Tag].Phase;
   			2:	Criteria2Tag := Criteria2Tag + PhaseNumber; (*Add phase number to address correct step totalizer*)
   				Criteria2RealValue := PhaseTotalizer[Criteria2Tag].Step;
   			3:	Criteria2RealValue := PhaseTotalizer[Criteria2Tag].Pause;
   			4:	Criteria2RealValue := PhaseTotalizer[Criteria2Tag].User;
   			5:	Criteria2RealValue := PhaseTotalizer[Criteria2Tag].Procedure;
   			8:	Criteria2RealValue := Totalizer[Criteria2Tag].Total;
   		ELSE 	CCPSystem.Error := 5;
   		END_CASE;
   	13:	CASE	Criteria2Property OF (*Valves*)
   			2:	Criteria2RealValue := Valve[Criteria2Tag].StatusWord;
   		ELSE 	CCPSystem.Error := 5;
   		END_CASE;
   	15:	CASE	Criteria2Property OF (*Misc.*)
   			1:	Criteria2BoolValue := MiscBOOL[Criteria2Tag];
   				Criteria2Type := 1;
   			2:	Criteria2RealValue := MiscDINT[Criteria2Tag];
   			3:	Criteria2RealValue := MiscREAL[Criteria2Tag];
   		ELSE 	CCPSystem.Error := 5;
   		END_CASE;
   	17:	CASE	Criteria2Property OF (*Miscellaneous*)
   			11:	Criteria2BoolValue := CCPSystem.DefaultOnComplete ;
   				Criteria2Type := 1;
   		ELSE 	CCPSystem.Error := 5;
   		END_CASE;
   	18:	CASE	Criteria2Property OF (*Criteria Flag*)
   			1:	Criteria2BoolValue := CriteriaFlag.Flag1 ;
   				Criteria2Type := 1;
   			2:	Criteria2BoolValue := CriteriaFlag.Flag2 ;
   				Criteria2Type := 1;
   			3:	Criteria2BoolValue := CriteriaFlag.Flag3 ;
   				Criteria2Type := 1;
   			4:	Criteria2BoolValue := CriteriaFlag.Flag4 ;
   				Criteria2Type := 1;
   			5:	Criteria2BoolValue := CriteriaFlag.Flag5 ;
   				Criteria2Type := 1;
   		ELSE 	CCPSystem.Error := 5;
   		END_CASE;
   	19:	CASE	Criteria2Property OF (*Concentration*)
   			1:	Criteria2RealValue := Concentration.VCF;
   			2:	Criteria2RealValue := Concentration.CB;
   			3:	Criteria2BoolValue := Concentration.Final_Conc_Volume_Reached ;
   				Criteria2Type := 1;
   			4:	Criteria2BoolValue := Concentration.Final_Conc_Protein_Reached ;
   				Criteria2Type := 1;
   		ELSE 	CCPSystem.Error := 5;
   		END_CASE;
   	20:	CASE	Criteria2Property OF (*Diafiltration*)
   			1:	Criteria2RealValue := Diafiltration.Diaf_Volume;
   			2:	Criteria2BoolValue := Diafiltration.Final_Diaf_Volum_Reached ;
   				Criteria2Type := 1;
   		ELSE 	CCPSystem.Error := 5;
   		END_CASE;
   	25: 	CASE	Criteria2Property OF (*Flow Paths*)
   			2:	Criteria2BoolValue := FlowPath[Criteria2Tag].Status;
   				Criteria2Type := 1;
   		ELSE 	CCPSystem.Error := 5;
   		END_CASE;
   	30: CASE	Criteria2Tag OF (*DCS*)
   			0:	Criteria2BoolValue := DCS.Criteria.Criteria_1;
   				Criteria2Type := 1;
   			1:	Criteria2BoolValue := DCS.Criteria.Criteria_2;
   				Criteria2Type := 1;
   		ELSE 	CCPSystem.Error := 5;
   		END_CASE;
   ELSE	CCPSystem.Error := 5;
   END_CASE;
   
END_ROUTINE
